(* Logix 5000 project; controller TFF vendor 1 type 14 code 107 rev 33.11; software revision 33.04; part 18 of 38 *)
(* tags used below, declared in another part *)
   _150S1 : ALIAS FOR DigitalOutput[0];
   AlarmControl : AlarmControl;   // Alarm Control
   ALM001 : ALIAS FOR DigitalOutput[2];
   BAN002P : ALIAS FOR DigitalOutput[6];
   BAN002S : ALIAS FOR DigitalOutput[5];
   ControlLoop : ControlLoop[20];   // Control Loop Array
   ControlLoop_PCV101_5ms : ALIAS FOR ControlLoop[4];
   ControlLoop_PCV201 : ALIAS FOR ControlLoop[5];
   ControlLoop_PCV201_5ms : ALIAS FOR ControlLoop[6];
   ControlLoop_PCV201Alarm : ALIAS FOR AlarmDeviation[5];
   CPU_Scanning : BOOL;   // System Scanning Flag
   ES001 : ALIAS FOR DigitalPoint[2];
   FirstScanComplete : BOOL;   // First Scan Complete Flag
   LI101 : ALIAS FOR AnalogPoint[44];
   Membrane_Data : Membrane_Data;   // Membrane Data
   Options : Options;   // Options List
   PCV101 : ALIAS FOR AnalogPoint[3];
   PCV201 : ALIAS FOR AnalogPoint[4];
   PCV201_AO : ALIAS FOR AnalogOutput[4];
   PCV201_Control : PCV_Control;   // PCV201 Control UDT
   PCV201_CVTune : CVTune;
   PCV201_PID : PCV;   // PCV201 PID Management
   Phase0 : ALIAS FOR Phase[0];   // Phase 0
   PLCFault : FaultRecordType;   // PLC Major Fault Record
   Rack_ACT350_WI101_200L : IO_Station;   // Status of ACT350 200L
   Rack_ACT350_WI101_500L : IO_Station;   // Status of ACT350 500L
   Rack_Murr_Node1_TFF20 : IO_Station;   // Status of Node 1 TFF20
   Rack_Murr_Node1_TFF40 : IO_Station;   // Status of Node 1 TFF40
   Rack_Murr_Node1_TFF80 : IO_Station;   // Status of Node 1 TFF80
   RawAnalogInputArray : INT[50];   // Array of analog input raw
   RSBUZZ : ALIAS FOR DigitalPoint[3];
   ScaleFiltering : ScaleFiltering;   // Data for Scale Filtering
   SysControl : SysControl;   // General system status and command
   ThisSystem : SystemType;
   TMP : ALIAS FOR AnalogPoint[41];
   Valve : Valve[100];   // Valve Array
   ValveControl : ValveControl;   // Valve Control
   WI101 : ALIAS FOR AnalogPoint[15];
   WI101Alarm : ALIAS FOR AlarmAnalog[15];
   WI201 : ALIAS FOR AnalogPoint[1];
   WI201Alarm : ALIAS FOR AlarmAnalog[1];
   YA10 : ALIAS FOR DigitalPoint[59];
(* MainProgram5ms, continued *)

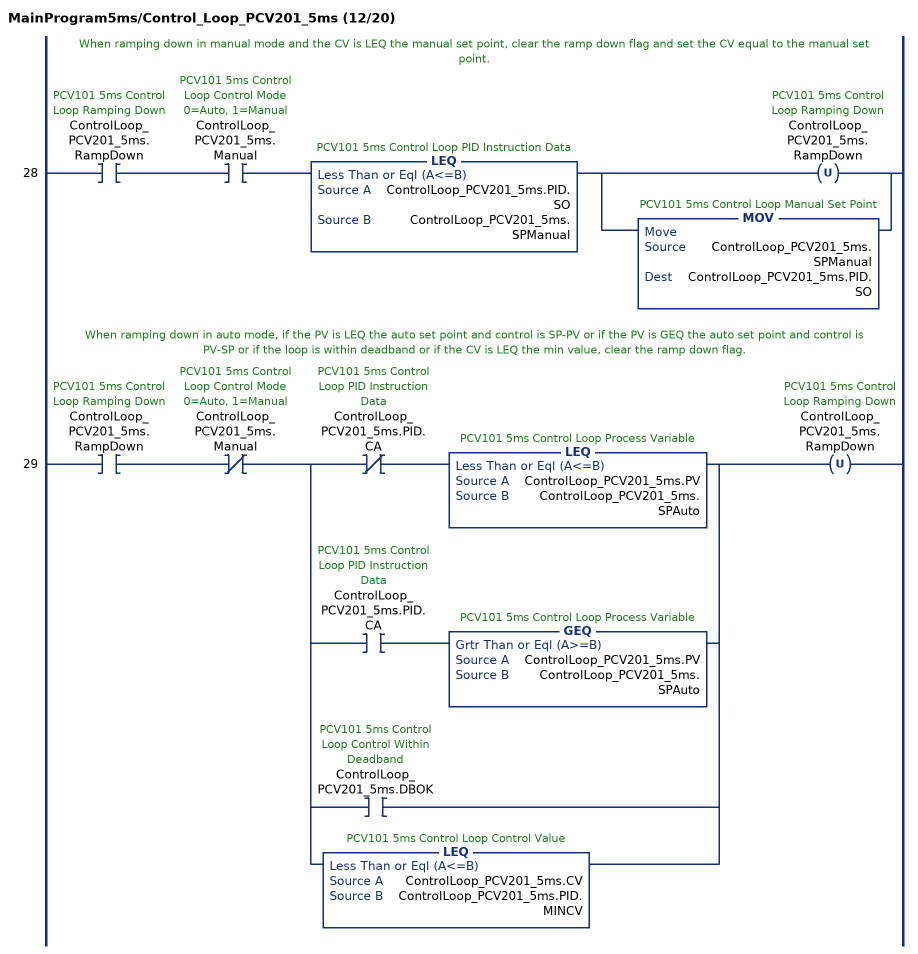
   // When ramping down in manual mode and the CV is LEQ the manual set point, clear the ramp down flag and set the CV equal to the manual set point.
   28: XIC(ControlLoop_PCV201_5ms.RampDown)XIC(ControlLoop_PCV201_5ms.Manual)LEQ(ControlLoop_PCV201_5ms.PID.SO,ControlLoop_PCV201_5ms.SPManual)[OTU(ControlLoop_PCV201_5ms.RampDown) ,MOV(ControlLoop_PCV201_5ms.SPManual,ControlLoop_PCV201_5ms.PID.SO) ];
   // When ramping down in auto mode, if the PV is LEQ the auto set point and control is SP-PV or if the PV is GEQ the auto set point and control is PV-SP or if the loop is within deadband or if the CV is LEQ the min value, clear the ramp down flag.
   29: XIC(ControlLoop_PCV201_5ms.RampDown)XIO(ControlLoop_PCV201_5ms.Manual)[XIO(ControlLoop_PCV201_5ms.PID.CA) LEQ(ControlLoop_PCV201_5ms.PV,ControlLoop_PCV201_5ms.SPAuto) ,XIC(ControlLoop_PCV201_5ms.PID.CA) GEQ(ControlLoop_PCV201_5ms.PV,ControlLoop_PCV201_5ms.SPAuto) ,XIC(ControlLoop_PCV201_5ms.DBOK) ,LEQ(ControlLoop_PCV201_5ms.CV,ControlLoop_PCV201_5ms.PID.MINCV) ]OTU(ControlLoop_PCV201_5ms.RampDown);
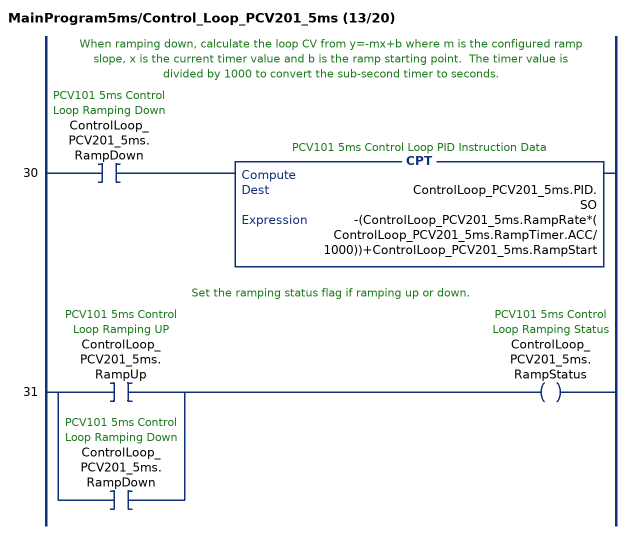
   // When ramping down, calculate the loop CV from y=-mx+b where m is the configured ramp slope, x is the current timer value and b is the ramp starting point.  The timer value is divided by 1000 to convert the sub-second timer to seconds.
   30: XIC(ControlLoop_PCV201_5ms.RampDown)CPT(ControlLoop_PCV201_5ms.PID.SO,-(ControlLoop_PCV201_5ms.RampRate*(ControlLoop_PCV201_5ms.RampTimer.ACC/1000))+ControlLoop_PCV201_5ms.RampStart);
   // Set the ramping status flag if ramping up or down.
   31: [XIC(ControlLoop_PCV201_5ms.RampUp) ,XIC(ControlLoop_PCV201_5ms.RampDown) ]OTE(ControlLoop_PCV201_5ms.RampStatus);
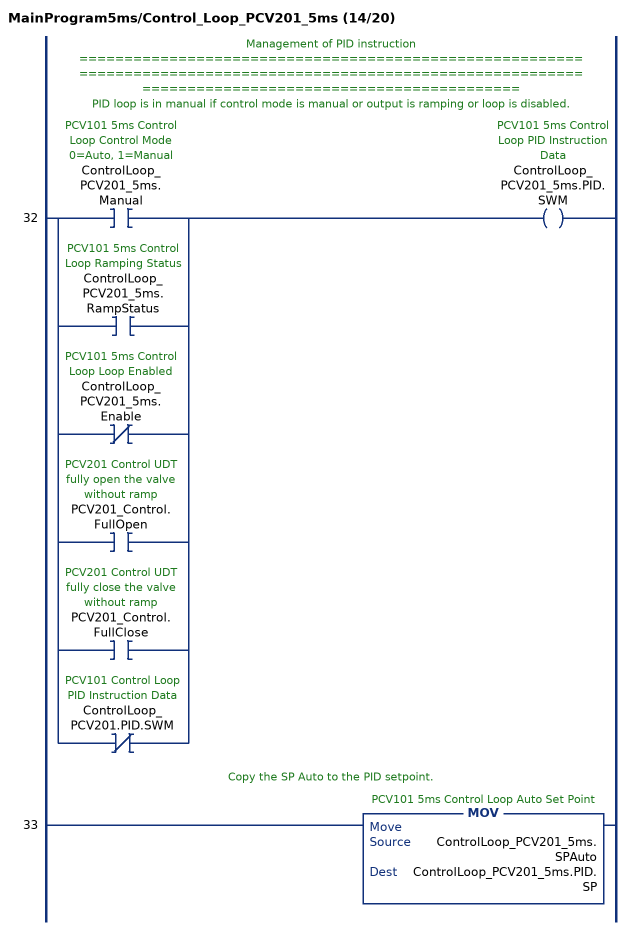
   // Management of PID instruction
   // ==========================================================================================================================================================
   // PID loop is in manual if control mode is manual or output is ramping or loop is disabled.
   32: [XIC(ControlLoop_PCV201_5ms.Manual) ,XIC(ControlLoop_PCV201_5ms.RampStatus) ,XIO(ControlLoop_PCV201_5ms.Enable) ,[[XIC(PCV201_Control.FullOpen) ,XIC(PCV201_Control.FullClose) ] ,XIO(ControlLoop_PCV201.PID.SWM) ] ]OTE(ControlLoop_PCV201_5ms.PID.SWM);
   // Copy the SP Auto to the PID setpoint.
   33: MOV(ControlLoop_PCV201_5ms.SPAuto,ControlLoop_PCV201_5ms.PID.SP);
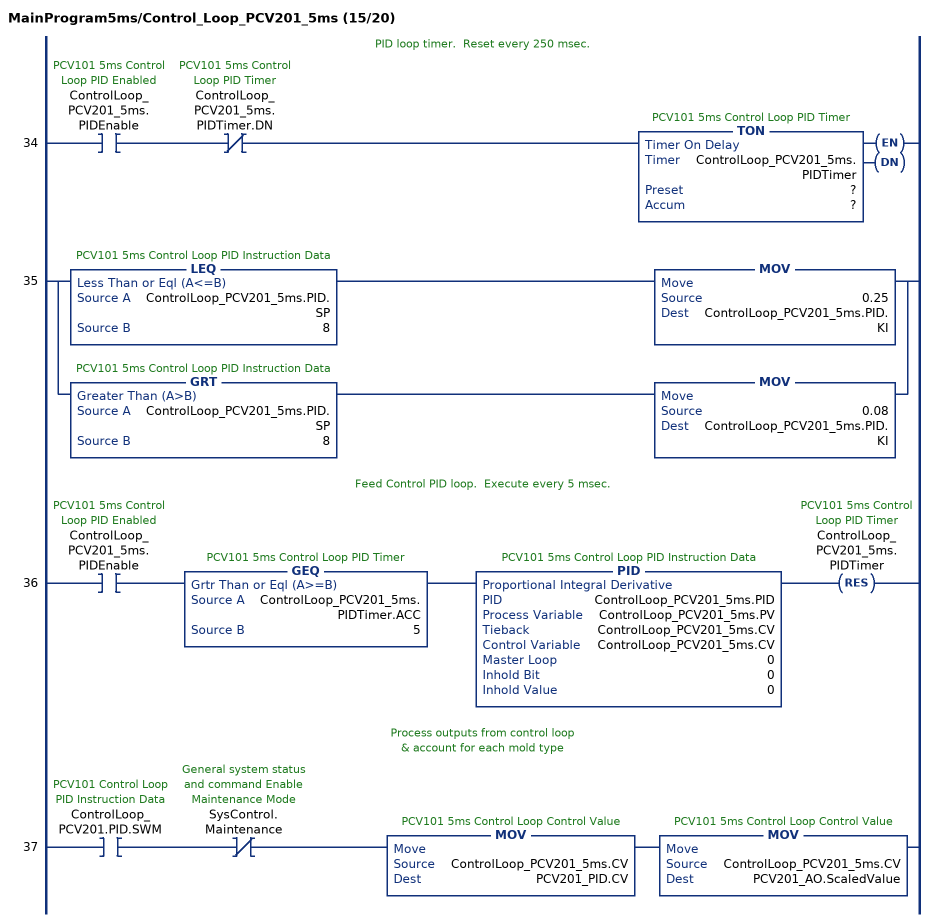
   // PID loop timer.  Reset every 250 msec.
   34: XIC(ControlLoop_PCV201_5ms.PIDEnable)XIO(ControlLoop_PCV201_5ms.PIDTimer.DN)TON(ControlLoop_PCV201_5ms.PIDTimer,?,?);
   35: [LEQ(ControlLoop_PCV201_5ms.PID.SP,8) MOV(0.25,ControlLoop_PCV201_5ms.PID.KI) ,GRT(ControlLoop_PCV201_5ms.PID.SP,8) MOV(0.08,ControlLoop_PCV201_5ms.PID.KI) ];
   // Feed Control PID loop.  Execute every 5 msec.
   36: XIC(ControlLoop_PCV201_5ms.PIDEnable)GEQ(ControlLoop_PCV201_5ms.PIDTimer.ACC,5)PID(ControlLoop_PCV201_5ms.PID,ControlLoop_PCV201_5ms.PV,ControlLoop_PCV201_5ms.CV,ControlLoop_PCV201_5ms.CV,0,0,0)RES(ControlLoop_PCV201_5ms.PIDTimer);
   // Process outputs from control loop
   // & account for each mold type
   37: XIC(ControlLoop_PCV201.PID.SWM)XIO(SysControl.Maintenance)MOV(ControlLoop_PCV201_5ms.CV,PCV201_PID.CV)MOV(ControlLoop_PCV201_5ms.CV,PCV201_AO.ScaledValue);
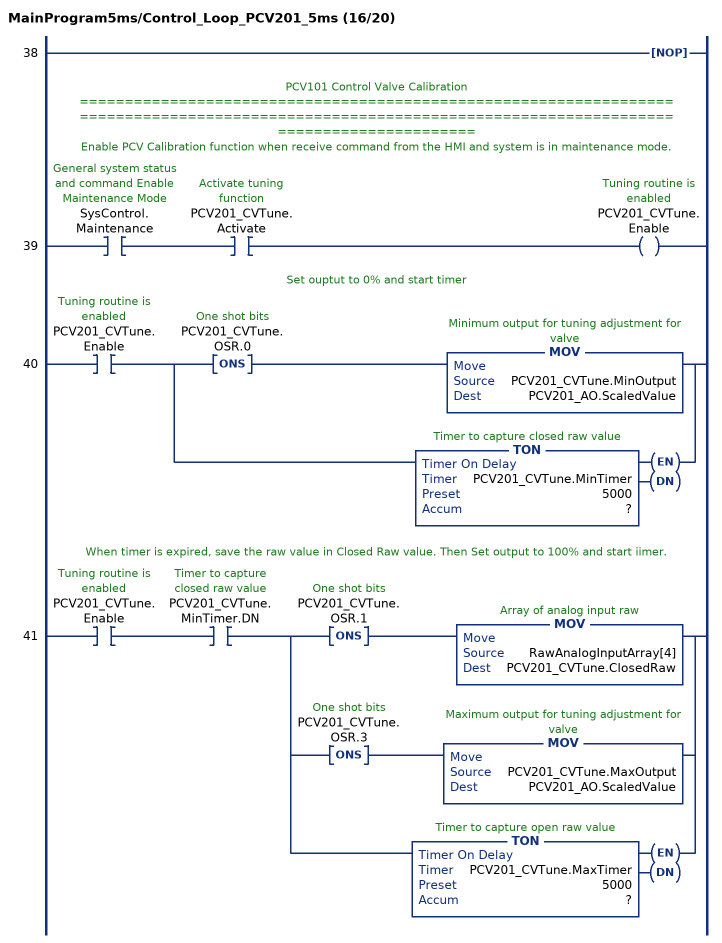
   38: NOP();
   // PCV101 Control Valve Calibration
   // ==========================================================================================================================================================
   // Enable PCV Calibration function when receive command from the HMI and system is in maintenance mode.
   39: XIC(SysControl.Maintenance)XIC(PCV201_CVTune.Activate)OTE(PCV201_CVTune.Enable);
   // Set ouptut to 0% and start timer
   40: XIC(PCV201_CVTune.Enable)[ONS(PCV201_CVTune.OSR.0) MOV(PCV201_CVTune.MinOutput,PCV201_AO.ScaledValue) ,TON(PCV201_CVTune.MinTimer,?,?) ];
   // When timer is expired, save the raw value in Closed Raw value. Then Set output to 100% and start iimer.
   41: XIC(PCV201_CVTune.Enable)XIC(PCV201_CVTune.MinTimer.DN)[ONS(PCV201_CVTune.OSR.1) MOV(RawAnalogInputArray[4],PCV201_CVTune.ClosedRaw) ,ONS(PCV201_CVTune.OSR.3) MOV(PCV201_CVTune.MaxOutput,PCV201_AO.ScaledValue) ,TON(PCV201_CVTune.MaxTimer,?,?) ];
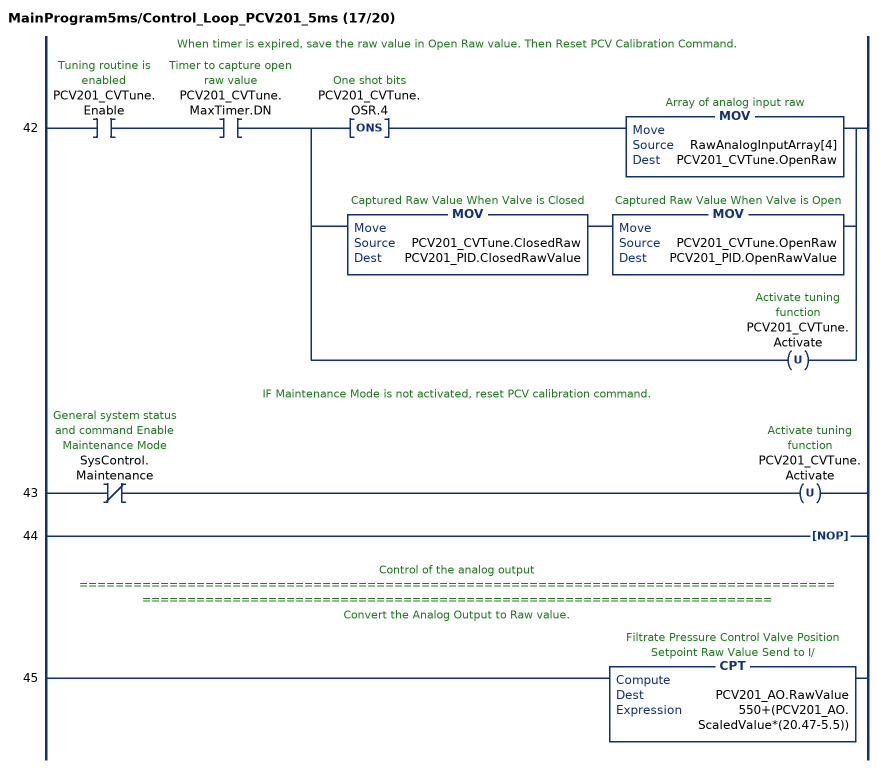
   // When timer is expired, save the raw value in Open Raw value. Then Reset PCV Calibration Command.
   42: XIC(PCV201_CVTune.Enable)XIC(PCV201_CVTune.MaxTimer.DN)[ONS(PCV201_CVTune.OSR.4) MOV(RawAnalogInputArray[4],PCV201_CVTune.OpenRaw) ,MOV(PCV201_CVTune.ClosedRaw,PCV201_PID.ClosedRawValue) MOV(PCV201_CVTune.OpenRaw,PCV201_PID.OpenRawValue) ,OTU(PCV201_CVTune.Activate) ];
   // IF Maintenance Mode is not activated, reset PCV calibration command.
   43: XIO(SysControl.Maintenance)OTU(PCV201_CVTune.Activate);
   44: NOP();
   // Control of the analog output
   // ==========================================================================================================================================================
   // Convert the Analog Output to Raw value.
   45: CPT(PCV201_AO.RawValue,550+(PCV201_AO.ScaledValue*(20.47-5.5)));
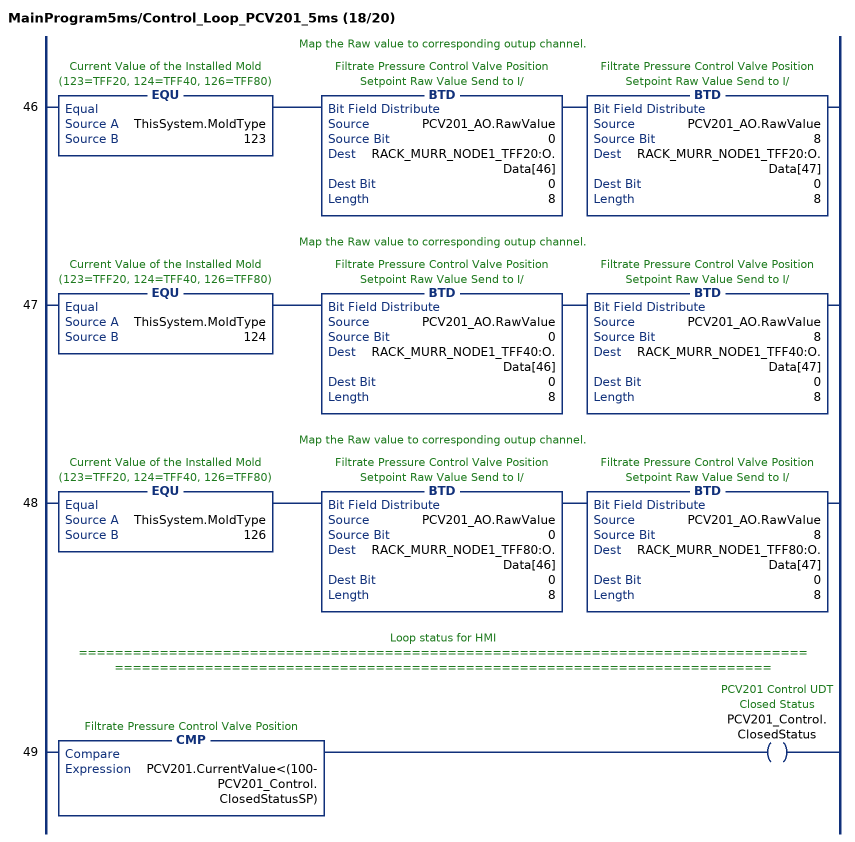
   // Map the Raw value to corresponding outup channel.
   46: EQU(ThisSystem.MoldType,123)BTD(PCV201_AO.RawValue,0,RACK_MURR_NODE1_TFF20:O.Data[46],0,8)BTD(PCV201_AO.RawValue,8,RACK_MURR_NODE1_TFF20:O.Data[47],0,8);
   // Map the Raw value to corresponding outup channel.
   47: EQU(ThisSystem.MoldType,124)BTD(PCV201_AO.RawValue,0,RACK_MURR_NODE1_TFF40:O.Data[46],0,8)BTD(PCV201_AO.RawValue,8,RACK_MURR_NODE1_TFF40:O.Data[47],0,8);
   // Map the Raw value to corresponding outup channel.
   48: EQU(ThisSystem.MoldType,126)BTD(PCV201_AO.RawValue,0,RACK_MURR_NODE1_TFF80:O.Data[46],0,8)BTD(PCV201_AO.RawValue,8,RACK_MURR_NODE1_TFF80:O.Data[47],0,8);
   // Loop status for HMI
   // ==========================================================================================================================================================
   49: CMP(PCV201.CurrentValue<(100-PCV201_Control.ClosedStatusSP))OTE(PCV201_Control.ClosedStatus);
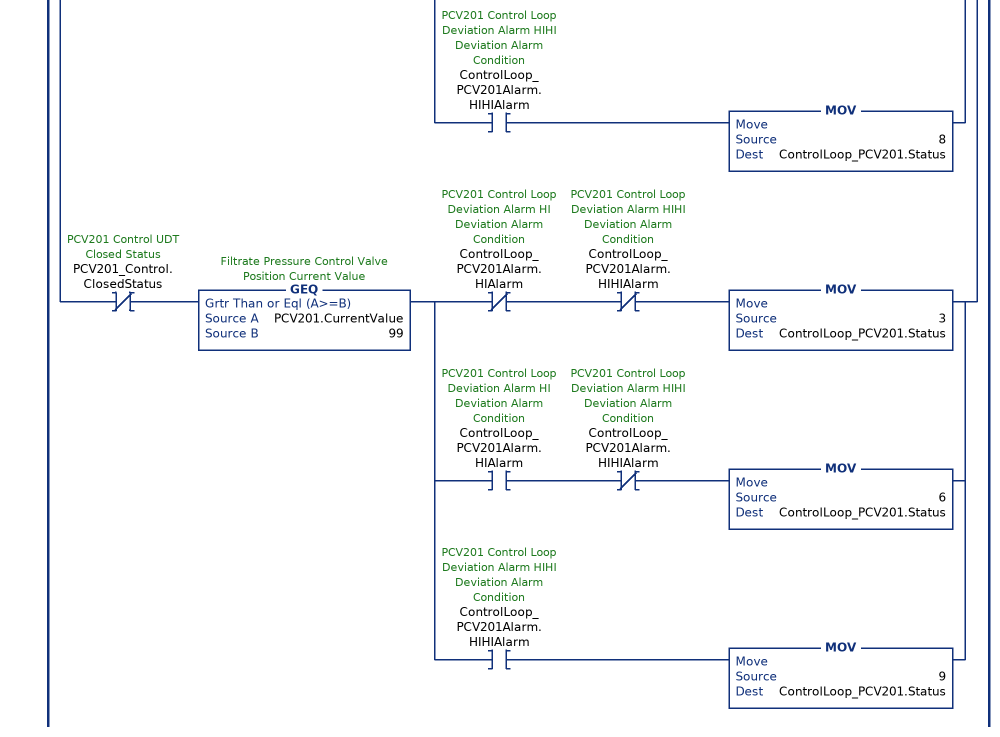
   // ControlLoop Status : 1 = PCV Close
   // ControlLoop Status : 2 = PCV Open
   // ControlLoop Status : 3 = PCV Full Open
   // ControlLoop Status : 4 = PCV Close and Non Critical alam
   // ControlLoop Status : 5 = PCV Open and Non Critical alam
   // ControlLoop Status : 6 = PCV Full Open and Non Critical alam
   // ControlLoop Status : 7 = PCV Close and Critical alam
   // ControlLoop Status : 8 = PCV Open and Critical alam
   // ControlLoop Status : 9 = PCV Full Open and Critical alam
   50: [XIC(PCV201_Control.ClosedStatus) [XIO(ControlLoop_PCV201Alarm.HIAlarm) XIO(ControlLoop_PCV201Alarm.HIHIAlarm) MOV(1,ControlLoop_PCV201.Status) ,XIC(ControlLoop_PCV201Alarm.HIAlarm) XIO(ControlLoop_PCV201Alarm.HIHIAlarm) MOV(4,ControlLoop_PCV201.Status) ,XIC(ControlLoop_PCV201Alarm.HIHIAlarm) MOV(7,ControlLoop_PCV201.Status) ] ,XIO(PCV201_Control.ClosedStatus) LES(PCV201.CurrentValue,99) [XIO(ControlLoop_PCV201Alarm.HIAlarm) XIO(ControlLoop_PCV201Alarm.HIHIAlarm) MOV(2,ControlLoop_PCV201.Status) ,XIC(ControlLoop_PCV201Alarm.HIAlarm) XIO(ControlLoop_PCV201Alarm.HIHIAlarm) MOV(5,ControlLoop_PCV201.Status) ,XIC(ControlLoop_PCV201Alarm.HIHIAlarm) MOV(8,ControlLoop_PCV201.Status) ] ,XIO(PCV201_Control.ClosedStatus) GEQ(PCV201.CurrentValue,99) [XIO(ControlLoop_PCV201Alarm.HIAlarm) XIO(ControlLoop_PCV201Alarm.HIHIAlarm) MOV(3,ControlLoop_PCV201.Status) ,XIC(ControlLoop_PCV201Alarm.HIAlarm) XIO(ControlLoop_PCV201Alarm.HIHIAlarm) MOV(6,ControlLoop_PCV201.Status) ,XIC(ControlLoop_PCV201Alarm.HIHIAlarm) MOV(9,ControlLoop_PCV201.Status) ] ];
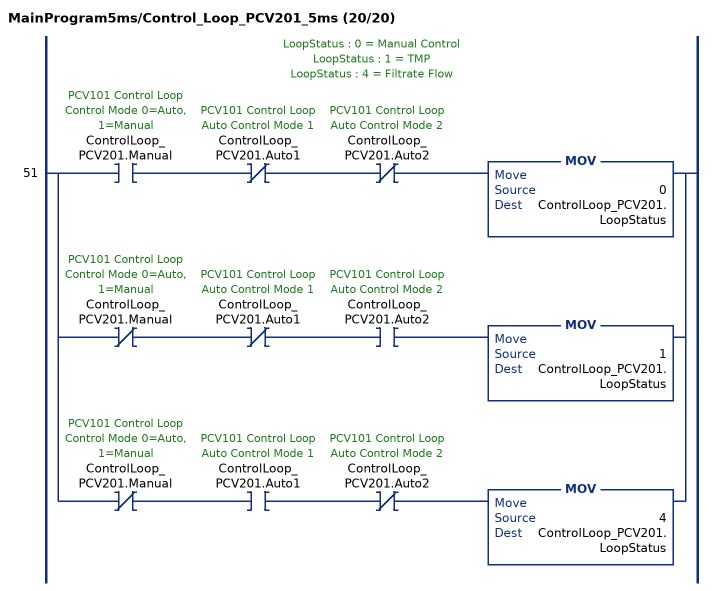
   // LoopStatus : 0 = Manual Control
   //  LoopStatus : 1 = TMP
   //  LoopStatus : 4 = Filtrate Flow
   51: [XIC(ControlLoop_PCV201.Manual) XIO(ControlLoop_PCV201.Auto1) XIO(ControlLoop_PCV201.Auto2) MOV(0,ControlLoop_PCV201.LoopStatus) ,XIO(ControlLoop_PCV201.Manual) XIO(ControlLoop_PCV201.Auto1) XIC(ControlLoop_PCV201.Auto2) MOV(1,ControlLoop_PCV201.LoopStatus) ,XIO(ControlLoop_PCV201.Manual) XIC(ControlLoop_PCV201.Auto1) XIO(ControlLoop_PCV201.Auto2) MOV(4,ControlLoop_PCV201.LoopStatus) ];
END_ROUTINE

ROUTINE FaultRoutine   (* ladder *)
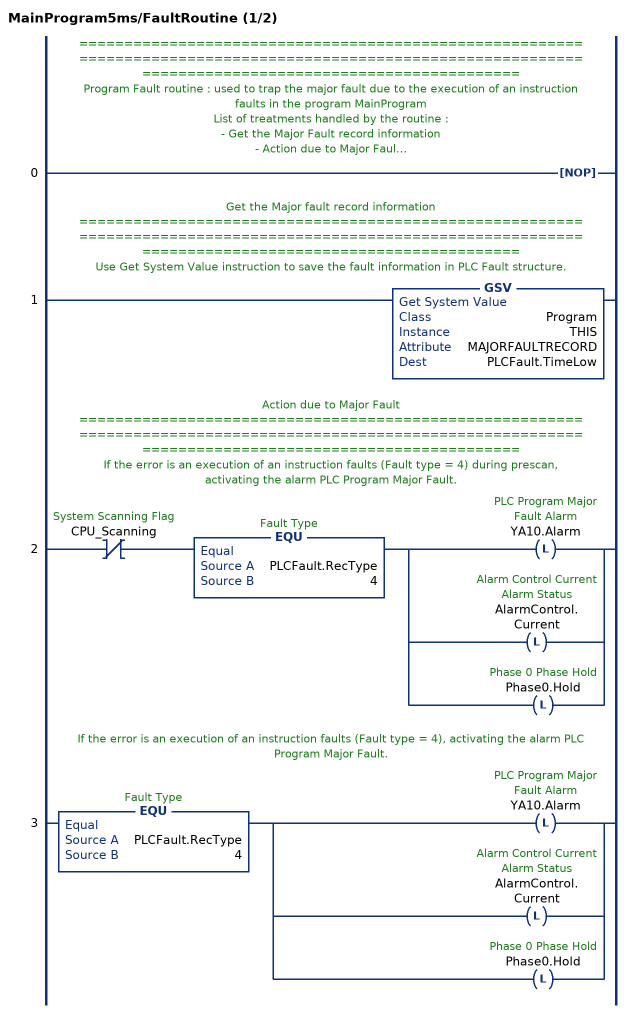
   // ==========================================================================================================================================================
   //                                                               Program Fault routine : used to trap the major fault due to the execution of an instruction faults in the program MainProgram
   //                                                     List of treatments handled by the routine :
   //                                                          - Get the Major Fault record information
   //                                                          - Action due to Major Fault
   //                                                     -----------------------------------------------------------------------------------------------------------------------------------------------------
   //                                                     History
   // 		2019-DEC-24 - Merck - Q. Spindler - Initial version for Candidate Release 1.00.00.00.a
   // ==========================================================================================================================================================
   0: NOP();
   // Get the Major fault record information
   // ==========================================================================================================================================================
   // Use Get System Value instruction to save the fault information in PLC Fault structure.
   1: GSV(Program,THIS,MAJORFAULTRECORD,PLCFault.TimeLow);
   // Action due to Major Fault
   // ==========================================================================================================================================================
   // If the error is an execution of an instruction faults (Fault type = 4) during prescan, activating the alarm PLC Program Major Fault.
   2: XIO(CPU_Scanning)EQU(PLCFault.RecType,4)[OTL(YA10.Alarm) ,OTL(AlarmControl.Current) ,OTL(Phase0.Hold) ];
   // If the error is an execution of an instruction faults (Fault type = 4), activating the alarm PLC Program Major Fault.
   3: EQU(PLCFault.RecType,4)[OTL(YA10.Alarm) ,OTL(AlarmControl.Current) ,OTL(Phase0.Hold) ];
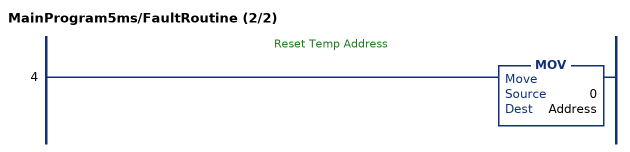
   // Reset Temp Address
   4: MOV(0,Address);
END_ROUTINE

ROUTINE Input_Analog_HighSpeed   (* ladder *)
// HighSpeed Analog Input Scaling
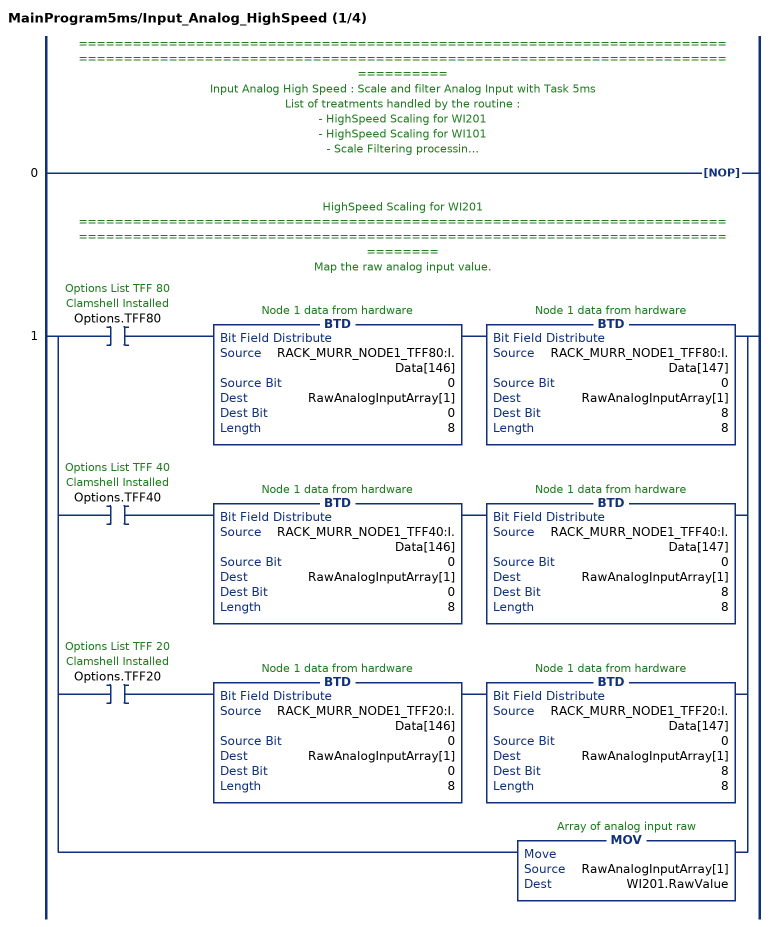
   // ==========================================================================================================================================================
   //                                                  Input Analog High Speed : Scale and filter Analog Input with Task 5ms
   //                                                     List of treatments handled by the routine :
   //                                                     - HighSpeed Scaling for WI201
   //                                                     - HighSpeed Scaling for WI101
   //                                                     - Scale Filtering processing
   //                                                     - Alarm Process Value Initialization
   //                                                     -----------------------------------------------------------------------------------------------------------------------------------------------------
   //                                                     History
   //      		2019-DEC-24 - Merck - Q. Spindler - Initial version for Candidate Release 1.00.00.00.a
   // ==========================================================================================================================================================
   0: NOP();
   // HighSpeed Scaling for WI201
   // ========================================================================================================================================================
   // Map the raw analog input value.
   1: [XIC(Options.TFF80) BTD(RACK_MURR_NODE1_TFF80:I.Data[146],0,RawAnalogInputArray[1],0,8) BTD(RACK_MURR_NODE1_TFF80:I.Data[147],0,RawAnalogInputArray[1],8,8) ,XIC(Options.TFF40) BTD(RACK_MURR_NODE1_TFF40:I.Data[146],0,RawAnalogInputArray[1],0,8) BTD(RACK_MURR_NODE1_TFF40:I.Data[147],0,RawAnalogInputArray[1],8,8) ,XIC(Options.TFF20) BTD(RACK_MURR_NODE1_TFF20:I.Data[146],0,RawAnalogInputArray[1],0,8) BTD(RACK_MURR_NODE1_TFF20:I.Data[147],0,RawAnalogInputArray[1],8,8) ,MOV(RawAnalogInputArray[1],WI201.RawValue) ];
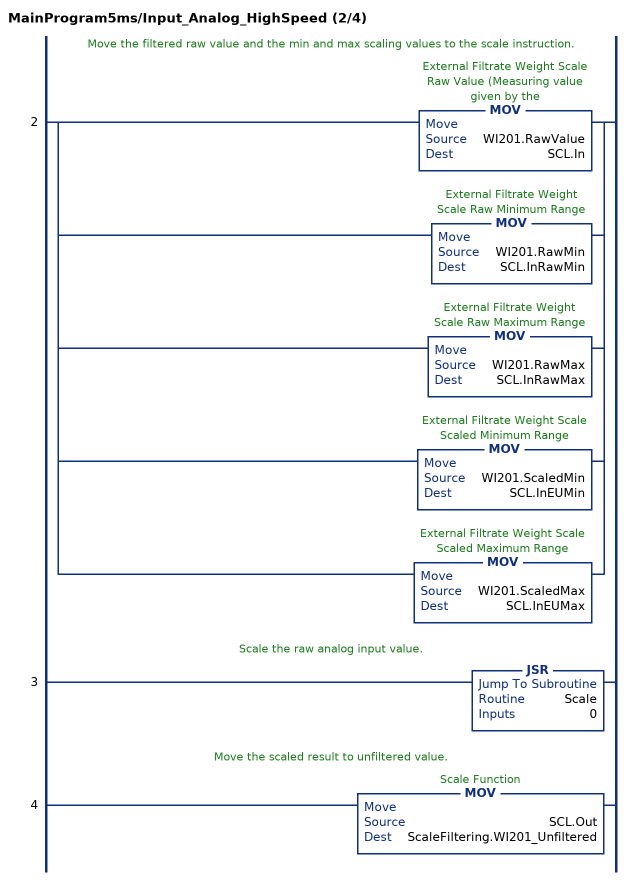
   // Move the filtered raw value and the min and max scaling values to the scale instruction.
   2: [MOV(WI201.RawValue,SCL.In) ,MOV(WI201.RawMin,SCL.InRawMin) ,MOV(WI201.RawMax,SCL.InRawMax) ,MOV(WI201.ScaledMin,SCL.InEUMin) ,MOV(WI201.ScaledMax,SCL.InEUMax) ];
   // Scale the raw analog input value.
   3: JSR(Scale,0);
   // Move the scaled result to unfiltered value.
   4: MOV(SCL.Out,ScaleFiltering.WI201_Unfiltered);
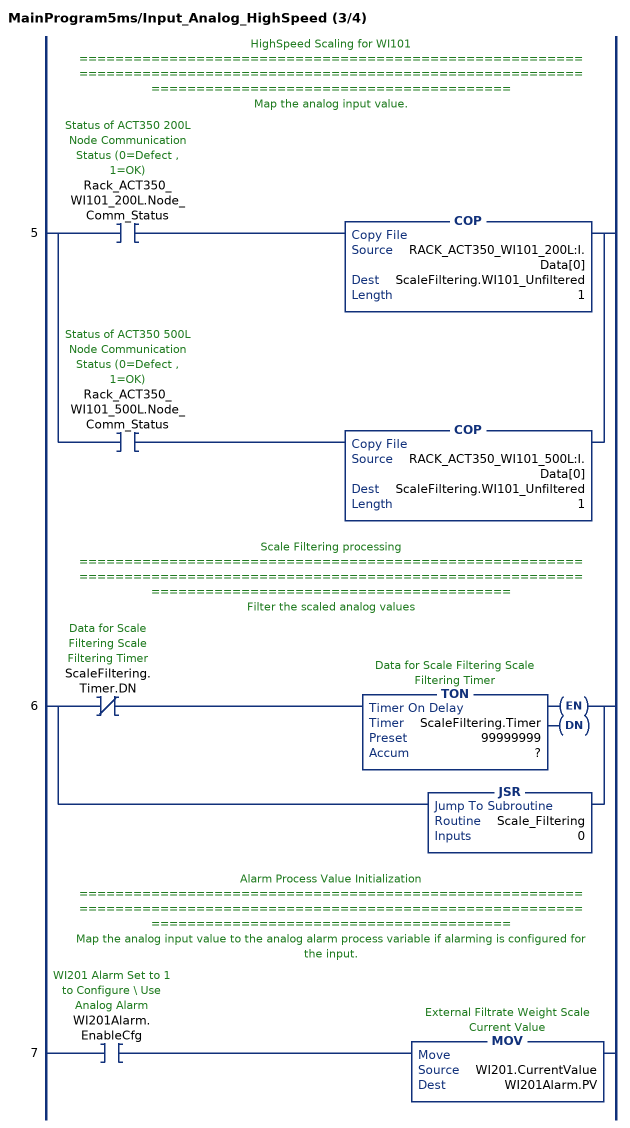
   // HighSpeed Scaling for WI101
   // ========================================================================================================================================================
   // Map the analog input value.
   5: [XIC(Rack_ACT350_WI101_200L.Node_Comm_Status) COP(RACK_ACT350_WI101_200L:I.Data[0],ScaleFiltering.WI101_Unfiltered,1) ,XIC(Rack_ACT350_WI101_500L.Node_Comm_Status) COP(RACK_ACT350_WI101_500L:I.Data[0],ScaleFiltering.WI101_Unfiltered,1) ];
   // Scale Filtering processing
   // ========================================================================================================================================================
   // Filter the scaled analog values
   6: [XIO(ScaleFiltering.Timer.DN) TON(ScaleFiltering.Timer,?,?) ,JSR(Scale_Filtering,0) ];
   // Alarm Process Value Initialization
   // ========================================================================================================================================================
   // Map the analog input value to the analog alarm process variable if alarming is configured for the input.
   7: XIC(WI201Alarm.EnableCfg)MOV(WI201.CurrentValue,WI201Alarm.PV);
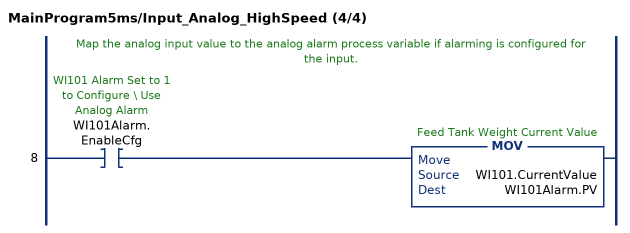
   // Map the analog input value to the analog alarm process variable if alarming is configured for the input.
   8: XIC(WI101Alarm.EnableCfg)MOV(WI101.CurrentValue,WI101Alarm.PV);
END_ROUTINE

ROUTINE MainRoutine   (* ladder *)
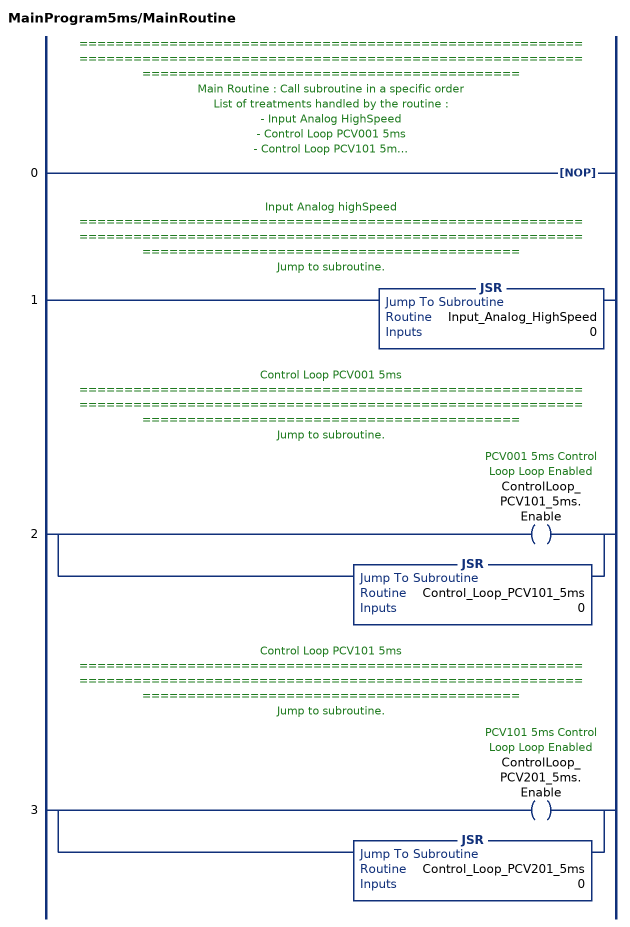
   // ==========================================================================================================================================================
   //                                                  Main Routine : Call subroutine in a specific order
   //                                                     List of treatments handled by the routine :
   //                                                - Input Analog HighSpeed
   //                                                - Control Loop PCV001 5ms
   //                                                - Control Loop PCV101 5ms
   //                                                     -----------------------------------------------------------------------------------------------------------------------------------------------------
   //                                                     History
   // 		2019-DEC-24 - Merck - Q. Spindler - Initial version for Candidate Release 1.00.00.00.a
   // ==========================================================================================================================================================
   0: NOP();
   // Input Analog highSpeed
   // ==========================================================================================================================================================
   // Jump to subroutine.
   1: JSR(Input_Analog_HighSpeed,0);
   // Control Loop PCV001 5ms
   // ==========================================================================================================================================================
   // Jump to subroutine.
   2: [OTE(ControlLoop_PCV101_5ms.Enable) ,JSR(Control_Loop_PCV101_5ms,0) ];
   // Control Loop PCV101 5ms
   // ==========================================================================================================================================================
   // Jump to subroutine.
   3: [OTE(ControlLoop_PCV201_5ms.Enable) ,JSR(Control_Loop_PCV201_5ms,0) ];
END_ROUTINE

ROUTINE Scale   (* function block diagram *)
// Scale Routine
   SHEET 1
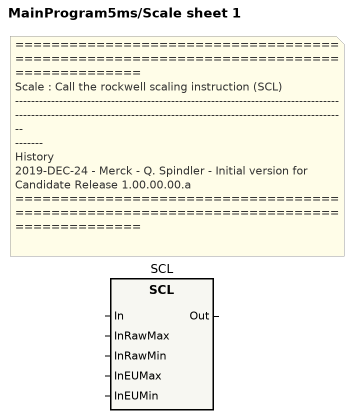
   // ======================================================================================
   // Scale : Call the rockwell scaling instruction (SCL)
   // --------------------------------------------------------------------------------------------------------------------------------------------------------------------
   // -------
   // History
   // 	2019-DEC-24 - Merck - Q. Spindler - Initial version for Candidate Release 1.00.00.00.a
   // ======================================================================================
   SCL : SCL();   // unwired pins: In InRawMax InRawMin InEUMax InEUMin Out
END_ROUTINE

ROUTINE Scale_Filtering   (* structured text *)
   
   (* =======================================================================
   	Scale Filtering : calculations of Filtered value
   
   	List of treatments
   		- Initialize Volume
   		- WI101 Feed Bag Volume Calculation
   		- Moving Average Filtering for Filtrate Volume
   		- Exponential Filtering for Filtrate Volume
   		- Analog Input processing
   
   -----------------------------------------------------------------------------------------------------------------------------------------------------
   	History
   		2019-DEC-24 - Merck - Q. Spindler - Initial version for Candidate Release 1.00.00.00.a
   =============================================================================================================================*)
   
   
   
   (* Initialize Volume
   =============================================================================================================================*)
   
   // Compute Volume values based on Unfiltered Weight and Density
   ScaleFiltering.FeedBagVolume := ScaleFiltering.WI101_Unfiltered / Membrane_Data.Density;
   ScaleFiltering.FiltrateVolume := ScaleFiltering.WI201_Unfiltered / Membrane_Data.Density;
   
   
   //Check that the minimum sample rate have met
   If ScaleFiltering.Timer.ACC > ScaleFiltering.Sample_Rate Then
   
   (* WI101 Feed Bag Volume Calculation
   =============================================================================================================================*)
   
   		//Compute the feed bag volume and Weight using the moving average filter
   		ScaleFiltering.FeedBagVolume_MAVE.In := ScaleFiltering.FeedBagVolume;
   		MAVE(ScaleFiltering.FeedBagVolume_MAVE, ScaleFiltering.FeedBagVolume_Array);
   		If Not SysControl.Simulate Then
   			LI101.CurrentValue := ScaleFiltering.FeedBagVolume_MAVE.Out;
   			WI101.CurrentValue := ScaleFiltering.FeedBagVolume_MAVE.Out * Membrane_Data.Density;
   		Else
   			LI101.CurrentValue := WI101.CurrentValue / Membrane_Data.Density;
   		End_If;
   
   (* Moving Average Filtering for Filtrate Volume
   =============================================================================================================================*)
   
   		//Compute the Filtrate volume and Weight using the moving average filter
   		ScaleFiltering.FiltrateVolume_MAVE.In := ScaleFiltering.FiltrateVolume;
   		MAVE(ScaleFiltering.FiltrateVolume_MAVE, ScaleFiltering.FiltrateVolume_Array);
   		ScaleFiltering.FiltrateVolume_MaveFiltered := ScaleFiltering.FiltrateVolume_MAVE.Out;
   		ScaleFiltering.Weight_MaveFiltered := ScaleFiltering.FiltrateVolume_MAVE.Out * Membrane_Data.Density;
   
   
   (* Exponential Filtering for Filtrate Volume
   =============================================================================================================================*)
   
   	//Compute the Filtrate volume using the Exponential filter
   	ScaleFiltering.FiltrateVolume_ExpFiltered := (ScaleFiltering.FiltrateVolume_ExpConst * ScaleFiltering.FiltrateVolume_ExpFiltered) + ((1-ScaleFiltering.FiltrateVolume_ExpConst)*ScaleFiltering.FiltrateVolume);
   
   	//Compute the Filtrate Weight using the filtered volume and density parameter
   	ScaleFiltering.Weight_ExpFiltered := ScaleFiltering.FiltrateVolume_ExpFiltered * Membrane_Data.Density;
   
   
   
   (* Analog Input processing
   =============================================================================================================================*)
   	//Assign Value to corresponding input
   		If ScaleFiltering.CurrentFilter = 0 Then //No Filtering
   			If Not SysControl.Simulate Then
   				WI201.CurrentValue := ScaleFiltering.FiltrateVolume * Membrane_Data.Density;
   			End_If;
   		End_If;
   
   		If ScaleFiltering.CurrentFilter = 1 Then //Moving Average Filter Active
   			If Not SysControl.Simulate Then
   				WI201.CurrentValue := ScaleFiltering.Weight_MaveFiltered;
   			End_If;
   		End_If;
   
   		If ScaleFiltering.CurrentFilter = 2 Then //Exponential Linear Recursive Filter active
   			If Not SysControl.Simulate Then
   				WI201.CurrentValue := ScaleFiltering.Weight_ExpFiltered;
   			End_If;
   		End_If;
   
   
   	ScaleFiltering.Timer.ACC := 0;
   
   	End_If;
END_ROUTINE
END_PROGRAM

PROGRAM Process   (* main routine MainRoutine, fault routine FaultRoutine *)
VAR
   Address : DINT := 111;   // Temp Address
   Address2 : DINT := 41;   // Temp Address
   AddressPump1 : DINT := 1;   // Temp Address for Pump 1
   AddressPump2 : DINT := 2;   // Temp Address for Pump 2
   AlarmInhibit_Timer : TIMER := (PRE := 500, ACC := 500);
   BufferSteps0_Prev : STRING25 := '81';
   Config : Configuration := (IndexA0 := 25, IndexAP := 50, IndexDP := 150, IndexDr := 11, IndeXValve := 100, IndexReset := 150, IndexCL := 20, IndexFlowpath := 61, IndexIOMod := 8);   // Index Array used in configuration routines
   FeedBagLevel_PID_Settings : INT;   // Index
   FeedPump_PID_Settings : INT;   // Index
   Index : DINT := 25;   // Index
   Index2 : DINT;   // Index
   Index3 : DINT;   // Index
   index4 : DINT := -1;   // Index
   initial_distribute : FBD_BIT_FIELD_DISTRIBUTE := (Source := 409663, SourceBit := 11, Length := 20, Dest := 200);
   ModbusLogTimer : TIMER := (PRE := 2000, ACC := 1756, EN := 1, TT := 1);
   NewSystem : DINT := 126;
   PCV001_PID_Settings : INT;
   PCV101_PID_Settings : INT;
   RecipeStepLog_DateTime_Empty : STRING25;   // Empty String
   RecipeStepLog_DateTime_Log : STRING25 := '10/03/2025 11:34:25 ';   // Last Date Time Received from HMI
   RecipeStepLog_DateTime_Prev : STRING25 := '10/03/2025 11:34:25 ';
   RecipeStepLog_Timer : TIMER := (PRE := 15000, ACC := 342, EN := 1, TT := 1);   // RecipeStepLog WatchDog Timer
   result : DINT[2] := ([0] := 1759491700);
   SCL : SCALE := (Status := 16#0000_0003, InstructFault := 1, InRawRangeInv := 1);   // Scale Instruction
   Temp1 : DINT := 324289;
   TIME : DINT[2] := ([0] := -1782024255, [1] := 409663);
   TimeInMicroSeconds : LINT := 1759491700324289;
   TimeInSeconds : LINT := 1759491700;
   TimeInSecondsDINT : DINT := 1759491700;
END_VAR

ROUTINE Alarm   (* ladder *)
// Alarm Routine
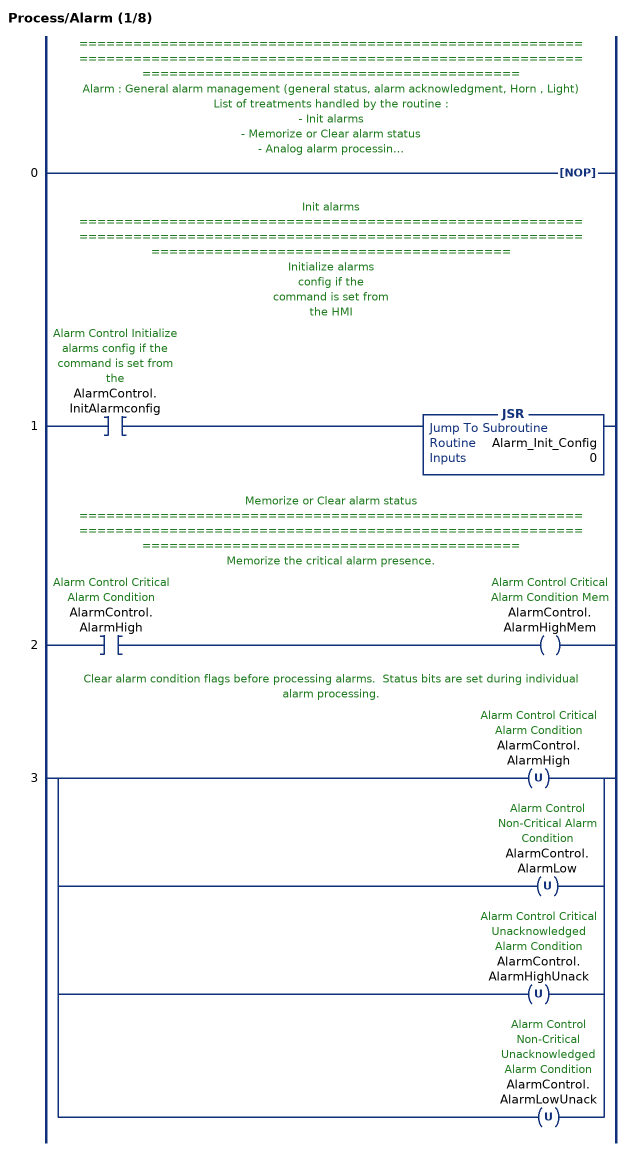
   // ==========================================================================================================================================================
   //                                                                                     Alarm : General alarm management (general status, alarm acknowledgment, Horn , Light)
   //                                                     List of treatments handled by the routine :
   //                                                         - Init alarms
   //                                                          - Memorize or Clear alarm status
   //                                                          - Analog alarm processing
   //                                                          - Deviation alarm processing
   //                                                          - Digital alarm processing
   //                                                          - General alarm status
   //                                                          - Flash control
   //                                                          - Alarm Horn
   //                                                          - Alarm Light
   //                                                          - Alarm acknowledgment
   //                                                          - Output processing
   //                                                     -----------------------------------------------------------------------------------------------------------------------------------------------------
   //                                                     History
   // 		2019-DEC-24 - Merck - Q. Spindler - Initial version for Candidate Release 1.00.00.00.a
   // 		2021-NOV-03 - Merck - Q. Spindler - Modifications for Candidate Release 1.01.00.00.a
   // - Add Init Alarms
   // ==========================================================================================================================================================
   0: NOP();
   // Init alarms
   // ========================================================================================================================================================
   //  Initialize alarms
   // config if the
   // command is set from
   // the HMI
   1: XIC(AlarmControl.InitAlarmconfig)JSR(Alarm_Init_Config,0);
   // Memorize or Clear alarm status
   // ==========================================================================================================================================================
   // Memorize the critical alarm presence.
   2: XIC(AlarmControl.AlarmHigh)OTE(AlarmControl.AlarmHighMem);
   // Clear alarm condition flags before processing alarms.  Status bits are set during individual alarm processing.
   3: [OTU(AlarmControl.AlarmHigh) ,OTU(AlarmControl.AlarmLow) ,OTU(AlarmControl.AlarmHighUnack) ,OTU(AlarmControl.AlarmLowUnack) ];
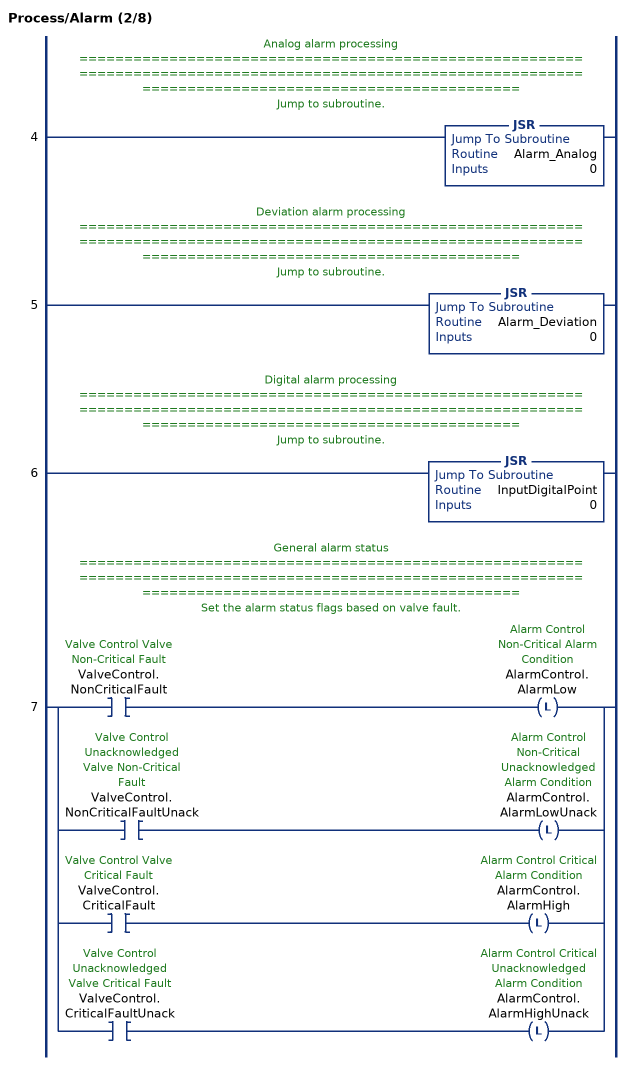
   // Analog alarm processing
   // ==========================================================================================================================================================
   // Jump to subroutine.
   4: JSR(Alarm_Analog,0);
   // Deviation alarm processing
   // ==========================================================================================================================================================
   // Jump to subroutine.
   5: JSR(Alarm_Deviation,0);
   // Digital alarm processing
   // ==========================================================================================================================================================
   // Jump to subroutine.
   6: JSR(InputDigitalPoint,0);
   // General alarm status
   // ==========================================================================================================================================================
   // Set the alarm status flags based on valve fault.
   7: [XIC(ValveControl.NonCriticalFault) OTL(AlarmControl.AlarmLow) ,XIC(ValveControl.NonCriticalFaultUnack) OTL(AlarmControl.AlarmLowUnack) ,XIC(ValveControl.CriticalFault) OTL(AlarmControl.AlarmHigh) ,XIC(ValveControl.CriticalFaultUnack) OTL(AlarmControl.AlarmHighUnack) ];
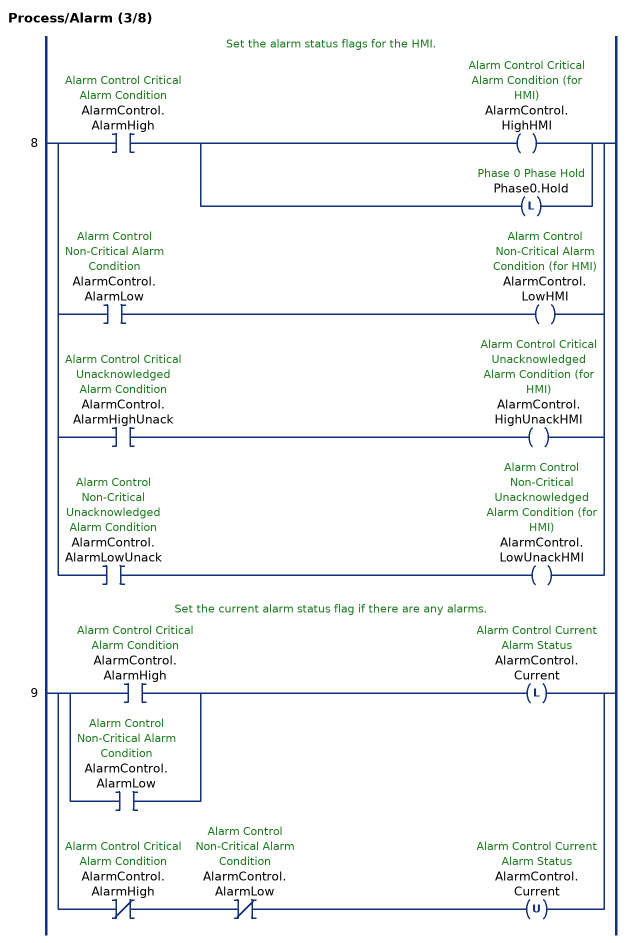
   // Set the alarm status flags for the HMI.
   8: [XIC(AlarmControl.AlarmHigh) [OTE(AlarmControl.HighHMI) ,OTL(Phase0.Hold) ] ,XIC(AlarmControl.AlarmLow) OTE(AlarmControl.LowHMI) ,XIC(AlarmControl.AlarmHighUnack) OTE(AlarmControl.HighUnackHMI) ,XIC(AlarmControl.AlarmLowUnack) OTE(AlarmControl.LowUnackHMI) ];
   // Set the current alarm status flag if there are any alarms.
   9: [[XIC(AlarmControl.AlarmHigh) ,XIC(AlarmControl.AlarmLow) ] OTL(AlarmControl.Current) ,XIO(AlarmControl.AlarmHigh) XIO(AlarmControl.AlarmLow) OTU(AlarmControl.Current) ];
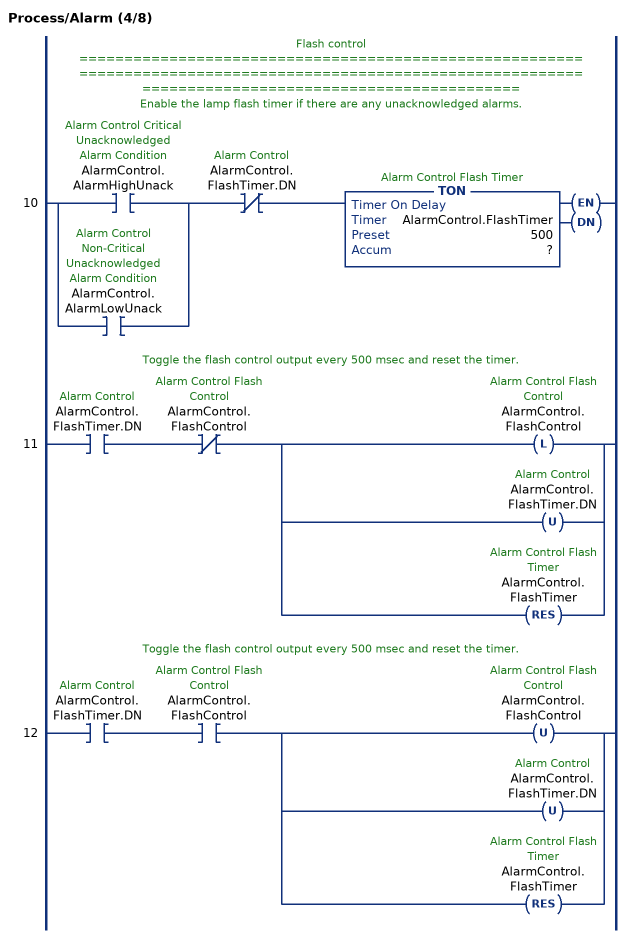
   // Flash control
   // ==========================================================================================================================================================
   // Enable the lamp flash timer if there are any unacknowledged alarms.
   10: [XIC(AlarmControl.AlarmHighUnack) ,XIC(AlarmControl.AlarmLowUnack) ]XIO(AlarmControl.FlashTimer.DN)TON(AlarmControl.FlashTimer,?,?);
   // Toggle the flash control output every 500 msec and reset the timer.
   11: XIC(AlarmControl.FlashTimer.DN)XIO(AlarmControl.FlashControl)[OTL(AlarmControl.FlashControl) ,OTU(AlarmControl.FlashTimer.DN) ,RES(AlarmControl.FlashTimer) ];
   // Toggle the flash control output every 500 msec and reset the timer.
   12: XIC(AlarmControl.FlashTimer.DN)XIC(AlarmControl.FlashControl)[OTU(AlarmControl.FlashControl) ,OTU(AlarmControl.FlashTimer.DN) ,RES(AlarmControl.FlashTimer) ];
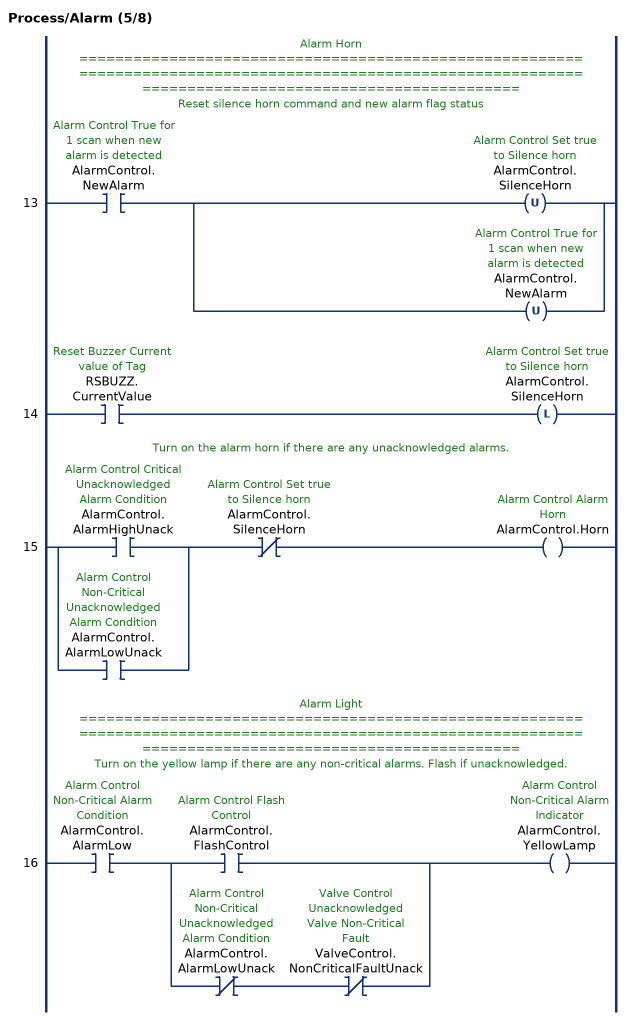
   // Alarm Horn
   // ==========================================================================================================================================================
   // Reset silence horn command and new alarm flag status
   13: XIC(AlarmControl.NewAlarm)[OTU(AlarmControl.SilenceHorn) ,OTU(AlarmControl.NewAlarm) ];
   14: XIC(RSBUZZ.CurrentValue)OTL(AlarmControl.SilenceHorn);
   // Turn on the alarm horn if there are any unacknowledged alarms.
   15: [XIC(AlarmControl.AlarmHighUnack) ,XIC(AlarmControl.AlarmLowUnack) ]XIO(AlarmControl.SilenceHorn)OTE(AlarmControl.Horn);
   // Alarm Light
   // ==========================================================================================================================================================
   // Turn on the yellow lamp if there are any non-critical alarms. Flash if unacknowledged.
   16: XIC(AlarmControl.AlarmLow)[XIC(AlarmControl.FlashControl) ,XIO(AlarmControl.AlarmLowUnack) XIO(ValveControl.NonCriticalFaultUnack) ]OTE(AlarmControl.YellowLamp);
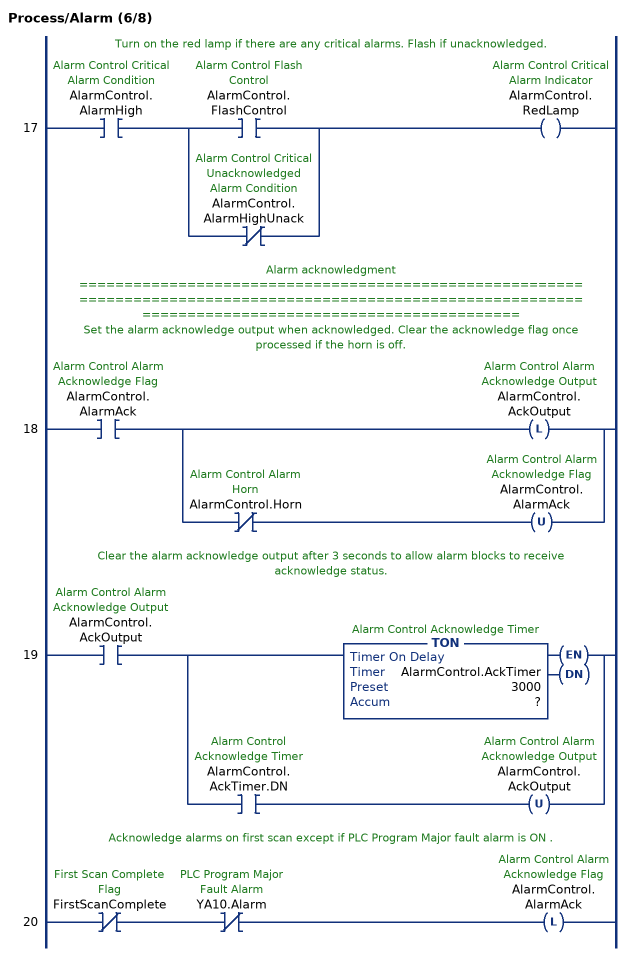
   // Turn on the red lamp if there are any critical alarms. Flash if unacknowledged.
   17: XIC(AlarmControl.AlarmHigh)[XIC(AlarmControl.FlashControl) ,XIO(AlarmControl.AlarmHighUnack) ]OTE(AlarmControl.RedLamp);
   // Alarm acknowledgment
   // ==========================================================================================================================================================
   // Set the alarm acknowledge output when acknowledged. Clear the acknowledge flag once processed if the horn is off.
   18: XIC(AlarmControl.AlarmAck)[OTL(AlarmControl.AckOutput) ,XIO(AlarmControl.Horn) OTU(AlarmControl.AlarmAck) ];
   // Clear the alarm acknowledge output after 3 seconds to allow alarm blocks to receive acknowledge status.
   19: XIC(AlarmControl.AckOutput)[TON(AlarmControl.AckTimer,?,?) ,XIC(AlarmControl.AckTimer.DN) OTU(AlarmControl.AckOutput) ];
   // Acknowledge alarms on first scan except if PLC Program Major fault alarm is ON .
   20: XIO(FirstScanComplete)XIO(YA10.Alarm)OTL(AlarmControl.AlarmAck);
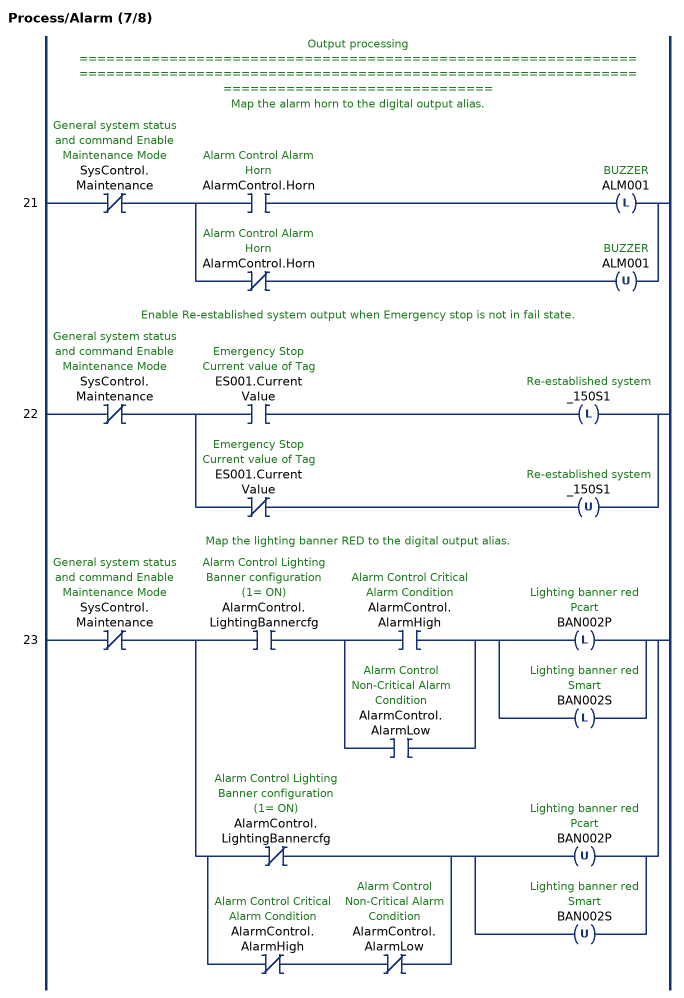
   // Output processing
   // ==========================================================================================================================================================
   // Map the alarm horn to the digital output alias.
   21: XIO(SysControl.Maintenance)[XIC(AlarmControl.Horn) OTL(ALM001) ,XIO(AlarmControl.Horn) OTU(ALM001) ];
   // Enable Re-established system output when Emergency stop is not in fail state.
   22: XIO(SysControl.Maintenance)[XIC(ES001.CurrentValue) OTL(_150S1) ,XIO(ES001.CurrentValue) OTU(_150S1) ];
   // Map the lighting banner RED to the digital output alias.
   23: XIO(SysControl.Maintenance)[XIC(AlarmControl.LightingBannercfg) [XIC(AlarmControl.AlarmHigh) ,XIC(AlarmControl.AlarmLow) ] [OTL(BAN002P) ,OTL(BAN002S) ] ,[XIO(AlarmControl.LightingBannercfg) ,XIO(AlarmControl.AlarmHigh) XIO(AlarmControl.AlarmLow) ] [OTU(BAN002P) ,OTU(BAN002S) ] ];
